(* PLC project , CODESYS CODESYS V3.5 SP16 Patch 4 *)
(* stored: creationDateTime 2021-05-04T13:17:28.6898035, modificationDateTime 2021-04-22T09:39:52.1420087 *)

PROGRAM th_X_trip
  VAR_INPUT
    f_X : INT;
  END_VAR
  VAR CONSTANT
    K_X_Min : INT := -55;
    k_X_Max : INT := 125;
  END_VAR
  VAR_INPUT
    f_Module_Error : BOOL;
    f_Channel_Error : BOOL;
    tx_X_Logic_Trip : BOOL;
  END_VAR
  VAR_OUTPUT
    tx_X_trip : BOOL;
  END_VAR

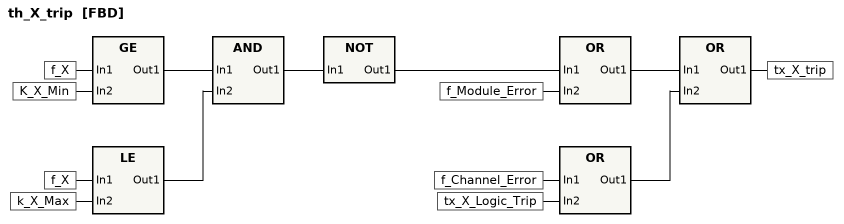
(* FBD diagram, written out as Structured Text *)
tx_X_trip := NOT (f_X >= K_X_Min AND f_X <= k_X_Max) OR f_Module_Error OR f_Channel_Error OR tx_X_Logic_Trip;
END_PROGRAM
